(* IEC 61131-3 sources: plc-vscode/tests/st/all/rusty/tests/lit/multi/constructors/src, 3 files *)

(* ---- main.st ---- *)
VAR_GLOBAL
    childInst : child;
END_VAR

FUNCTION main : DINT
    childInst();
    main := childInst.y + childInst.x; // Should be 36 (18 + 18)
    printf('%d$N', main);
END_FUNCTION

(* ---- base.st ---- *)
FUNCTION_BLOCK baseFb
    VAR_OUTPUT
        x : DINT;
        y : REFERENCE TO DINT REF= x;
    END_VAR

    METHOD FB_INIT
        THIS^.x := 10;
        THIS^.y := THIS^.x + 1; //x and y are 11
    END_METHOD
END_FUNCTION_BLOCK

(* ---- child.st ---- *)
FUNCTION_BLOCK child EXTENDS baseFb
    THIS^.x := This^.x + 5; // x is now 16
    THIS^.y := THIS^.y + 2; // y is now 18
END_FUNCTION_BLOCK
